// TIA Portal V21 export
FUNCTION_BLOCK "FB_AnaDoubleCall"   // FB12, SCL
TITLE = Analyzer: same instance called twice
{ S7_Optimized_Access := 'TRUE' }
// Rule C26b: the counter instance PartCounter is called twice in one cycle
// stored: MemoryReserve 100, SetENOAutomatically false
   VAR_INPUT
      PulseA : Bool;   // First count pulse
      PulseB : Bool;   // Second count pulse
   END_VAR
   VAR_OUTPUT
      Count : Int;   // Counter value
   END_VAR
   VAR
      PartCounter { S7_SetPoint := 'True'} : CTU_INT;   // Up counter
   END_VAR
BEGIN

       #PartCounter(CU := #PulseA, R := FALSE, PV := 100);
       #PartCounter(CU := #PulseB, R := FALSE, PV := 100);
       #Count := #PartCounter.CV;
END_FUNCTION_BLOCK
